DATA_BLOCK "World"
{ S7_Optimized_Access := 'TRUE' }
VERSION : 0.1
NON_RETAIN
   VAR
      Bay0 : Array[0..3, 0..11] of UInt;     // working copy of the ship (FB10 INIT copy / OB30 lift-put effect)
      Bay1 : Array[0..3, 0..11] of UInt;     // working copy of the yard
      CraneX : SInt;                         // crane x after last completed command
      CraneY : SInt;
      CraneBay : USInt := 1;
      Carried : UInt;                        // ID on the hook (0 = none)
      Busy : Bool;                           // command issued to FB1, not finished yet
      BusyTicks : Int;                       // OB30 ticks since issue (watchdog)
      ActCmd : "typeCmd";                    // command currently executing
      NextCmd : "typeCmd";                   // staged command (valid when CmdReady)
      CmdReady : Bool;                       // handshake: FB10 sets (last) / OB30 clears
      Permit : Bool;                         // OB30 may issue NextCmd
      DoneSeq : UDInt;                       // +1 per completed command
      LastDone : "typeCmd";                  // last completed command
      Fault : Word;                          // OB30-detected alarms (bit = alarm bit)
      FaultCmd : "typeCmd";                  // command rejected by CheckCmd
      UList : Array[1..48] of UInt;          // copy of DB20 (unload list)
      UState : Array[1..48] of USInt;        // 0 pending, 1 done, 2 skipped
      LList : Array[1..48] of UInt;          // copy of DB21 (load list)
      LState : Array[1..48] of USInt;        // as UState
      N : Int;                               // non-zero entries in DB20 + DB21 (for J)
      Plan : Array[1..96] of "typeTransfer"; // written by the planner
      PlanLen : Int;
      PlanValid : Bool;
      PlanVariant : Int;
      PredT_ds : DInt;
      PredM : DInt;
      PredJ : Real;
      BaseT_ds : DInt;                       // ROUND(T*10) at plan request
      BaseM : DInt;                          // M at plan request
      PlanIdx : Int := 1;                    // done pointer: transfer being executed
      Phase : USInt;                         // done pointer: next phase of PlanIdx to complete
      StageIdx : Int := 1;                   // staging cursor (transfer)
      StagePhase : USInt;                    // staging cursor (phase)
      BalL : Int;                            // ship count x in {0,1}
      BalR : Int;                            // ship count x in {2,3}
      BalF : Int;                            // ship count y in 0..5
      BalA : Int;                            // ship count y in 6..11
      CfgOrderMode : USInt := 1;             // 0 free, 1 per-list order, 2 strict (set by FB10 from HMI_IF before each plan)
      CfgBalLimit : Int := 5;
      CfgBalMode : USInt;                    // 0 x-halves only, 1 also y-halves
      CfgMMode : USInt := 0;                 // manipulation count model (CONTRACT 4.1); v1.7: 0 = spec rule (diagonal = 2), 2 = FB1 (+1 per move command)
      CfgVariants : Int := 4;
      CfgAlpha : Array[1..4] of Int := [0, 75, 125, 200];    // v1.7: retuned for CfgMMode 0 (v1.3 mode 2: [0, 100, 200, 300])
      CfgStepsPerCall : Int := 1;
      CfgTimeoutTicks : Int := 10;           // FB1 watchdog in OB30 ticks (1 s)
      OB30Ticks : UDInt;
      MSpec : UDInt;                         // manipulations by the spec rule (OB30): +1 per changed axis, +1 lift/put
      // ---- v1.3: improve phase (CONTRACT 4.8) and lower bound (4.9) ----
      CfgImproveEvals : DInt := 3000;        // local-search evaluations after the greedy (0 = off)
      CfgImproveDist : Int := 0;             // max |i-j| of a move (0 = unlimited)
      CfgImprovePerCall : Int := 1;          // evaluations per OB1 call (per-call work bound)
      PredJ0 : Real;                         // J of the greedy winner before the improve phase
      LbT_ds : DInt;                         // lower bound of the final T (incl. BaseT_ds), deciseconds
      LbM : DInt;                            // lower bound of the final M (incl. BaseM)
      LbJ : Real;                            // lower bound of J (no plan can be better)
      ImpEvals : DInt;                       // improve phase: evaluations done (last plan)
      ImpAccepts : DInt;                     // improve phase: accepted improvements (last plan)
      // ---- v1.4: exact order feasibility (CONTRACT 4.10) and SLOT phase (4.11) ----
      CfgSlotSweeps : Int := 10;             // drop-cell local search sweeps after IMPROVE (0 = off)
      SlotAccepts : DInt;                    // SLOT phase: accepted drop-cell changes (last plan)
      OrderFeasible : Bool;                  // last plan job: the requested order mode is feasible (exact DP)
      // ---- v1.5 (judge round 2 R2-J1): relaxed balance rule on a ship that starts out of balance ----
      BalCeil : Int;                         // 0 = step rule; > CfgBalLimit: while |L-R| > CfgBalLimit a step may go up to BalCeil
      // ---- v1.6 (judge round 3 R3-E3): relaxed ceiling search ----
      CfgRelaxMin : Bool;                    // FALSE: relaxed fallback uses BalCeil = start imbalance at once; TRUE: ascending CfgBalLimit+1 .. start imbalance (smallest feasible, costs J)
   END_VAR


BEGIN

END_DATA_BLOCK

